(* IEC 61131-3 sources: codesys-to-s7/tests/corpus/C2S7-POU-STAT/pos, 1 file *)

(* ---- input.st ---- *)
FUNCTION F_Case : INT
VAR_STAT
    n : INT;
END_VAR
n := n + 1; F_Case := n;
END_FUNCTION
